(* PLC project Claude3.project, CODESYS CODESYS V3.5 SP20 *)
(* stored: creationDateTime 2026-10-23T09:23:11.8560198, modificationDateTime 2026-10-23T09:22:48.4769723 *)

(* values of E_LineState: DISABLED: Linha desabilitada; WAIT_BOTTLE: Aguardando lote / garrafa; CLAMPING: Cilindro travando a garrafa + tara; FILLING: Enchendo; DRIPPING: Gotejamento, válvula fechada; UNCLAMPING: Cilindro liberando a garrafa; DONE: Ciclo concluído, aguarda avanço da esteira; FAULT: Falha travada, requer reset *)

{attribute 'qualified_only'}
{attribute 'strict'}
TYPE E_LineState : (DISABLED := 0, WAIT_BOTTLE := 1, CLAMPING := 2, FILLING := 3, DRIPPING := 4, UNCLAMPING := 5, DONE := 6, FAULT := 7);
END_TYPE

(* values of E_Fault: FILL_TIMEOUT: Tempo de enchimento excedido; CLAMP_TIMEOUT: Cilindro nao fechou no tempo; UNCLAMP_TIMEOUT: Cilindro nao abriu no tempo; BOTTLE_REMOVED: Garrafa removida durante o ciclo; SAFETY: Emergencia ou porta aberta *)

{attribute 'qualified_only'}
{attribute 'strict'}
TYPE E_Fault : (NONE := 0, FILL_TIMEOUT := 1, CLAMP_TIMEOUT := 2, UNCLAMP_TIMEOUT := 3, BOTTLE_REMOVED := 4, SAFETY := 5);
END_TYPE

(* values of E_ConvState: ADVANCE: Esteira avancando ate o proximo lote; SETTLE: Lote posicionado, tempo de acomodacao; PROCESSING: Linhas enchendo *)

{attribute 'qualified_only'}
{attribute 'strict'}
TYPE E_ConvState : (ADVANCE := 0, SETTLE := 1, PROCESSING := 2);
END_TYPE

TYPE ST_Recipe : STRUCT
  sName : STRING(20);  (* Nome da receita *)
  rTargetMass_g : REAL;  (* Massa liquida alvo [g] *)
  rPreAct_g : REAL;  (* Pre-atuacao: fecha a valvula antes do alvo [g] *)
  rTolerance_g : REAL;  (* Tolerancia +/- para aprovar a garrafa [g] *)
  tFillTimeout : TIME;  (* Tempo maximo de enchimento *)
  tDrip : TIME;  (* Tempo de gotejamento *)
END_STRUCT;
END_TYPE

FUNCTION_BLOCK FB_MovingAvg
  VAR_INPUT
    rIn : REAL;  (* Amostra atual *)
  END_VAR
  VAR_OUTPUT
    rOut : REAL;  (* Media das ultimas C_FILTER_SIZE amostras *)
  END_VAR
  VAR
    aBuf : ARRAY[0..(GVL_Main.C_FILTER_SIZE - 1)] OF REAL;
    iIdx : INT := 0;
    bInit : BOOL := FALSE;
    i : INT;
    rSum : REAL;
  END_VAR

                  (* Na primeira chamada, preenche o buffer para evitar transitorio *)
IF NOT bInit THEN
    FOR i := 0 TO GVL_Main.C_FILTER_SIZE - 1 DO
        aBuf[i] := rIn;
    END_FOR;
    bInit := TRUE;
END_IF;

(* Buffer circular *)
aBuf[iIdx] := rIn;
iIdx := iIdx + 1;
IF iIdx > GVL_Main.C_FILTER_SIZE - 1 THEN
    iIdx := 0;
END_IF;

(* Soma e media *)
rSum := 0.0;
FOR i := 0 TO GVL_Main.C_FILTER_SIZE - 1 DO
    rSum := rSum + aBuf[i];
END_FOR;
rOut := rSum / INT_TO_REAL(GVL_Main.C_FILTER_SIZE);
                
END_FUNCTION_BLOCK

FUNCTION_BLOCK FB_LevelControl
  VAR_INPUT
    bEnable : BOOL;  (* FALSE = fecha a valvula (seguranca) *)
    rLevel_pct : REAL;  (* Nivel atual [%] *)
    rLowOn_pct : REAL := 30.0;  (* Abre a valvula abaixo deste nivel *)
    rHighOff_pct : REAL := 80.0;  (* Fecha a valvula acima deste nivel *)
    rMinOperate_pct : REAL := 15.0;  (* Minimo para liberar o enchimento *)
  END_VAR
  VAR_OUTPUT
    bFillValve : BOOL;  (* Valvula de entrada do tanque *)
    bTankOk : BOOL;  (* Nivel suficiente para envasar *)
    bLowLevelAlarm : BOOL;
  END_VAR

                  (* Histerese: a saida mantem o ultimo estado entre os limites *)
IF NOT bEnable THEN
    bFillValve := FALSE;
ELSIF rLevel_pct <= rLowOn_pct THEN
    bFillValve := TRUE;
ELSIF rLevel_pct >= rHighOff_pct THEN
    bFillValve := FALSE;
END_IF;

(* Permissivo de envase e alarme de nivel baixo *)
bTankOk        := rLevel_pct >= rMinOperate_pct;
bLowLevelAlarm := NOT bTankOk;
                
END_FUNCTION_BLOCK

FUNCTION_BLOCK FB_FillLine
  VAR_INPUT
    bEnable : BOOL;  (* Linha habilitada *)
    bSafetyOk : BOOL;  (* Emergencia e porta OK *)
    bRun : BOOL;  (* Maquina em producao (permite iniciar garrafa) *)
    bLotReady : BOOL;  (* Lote posicionado e acomodado *)
    bTankOk : BOOL;  (* Nivel do tanque suficiente *)
    bBottlePresent : BOOL;
    bClampClosed : BOOL;
    bClampOpen : BOOL;
    bReset : BOOL;  (* Reset de falha (borda de subida) *)
    rMass_g : REAL;  (* Massa bruta filtrada *)
    stRecipe : ST_Recipe;
  END_VAR
  VAR_OUTPUT
    bClampCmd : BOOL;
    bFillValve : BOOL;
    bFinished : BOOL;  (* Desabilitada ou concluida no lote atual *)
    bBusy : BOOL;  (* Garrafa em processo *)
    bFault : BOOL;
    eState : E_LineState := E_LineState.DISABLED;
    eFault : E_Fault := E_Fault.NONE;
    rNetMass_g : REAL;
    diFilled : DINT;
    diRejected : DINT;
  END_VAR
  VAR
    trigReset : R_TRIG;
    tonClamp : TON;
    tonUnclamp : TON;
    tonTare : TON;
    tonFill : TON;
    tonDrip : TON;
    tonBottle : TON;
    rTare_g : REAL;
    bInProcess : BOOL;  (* Ha garrafa em processo nesta linha *)
    bFaultMidCycle : BOOL;  (* Falha ocorreu com garrafa em processo *)
    bWatchBottle : BOOL;
    eFaultNew : E_Fault;
  END_VAR

                  (* ---- 1. Temporizadores e deteccao de borda ---- *)
bWatchBottle := (eState = E_LineState.CLAMPING) OR (eState = E_LineState.FILLING)
                OR (eState = E_LineState.DRIPPING);

trigReset(CLK := bReset);
tonClamp  (IN := (eState = E_LineState.CLAMPING)   AND NOT bClampClosed, PT := GVL_Main.C_T_CYL_TIMEOUT);
tonTare   (IN := (eState = E_LineState.CLAMPING)   AND bClampClosed,     PT := GVL_Main.C_T_TARE);
tonUnclamp(IN := (eState = E_LineState.UNCLAMPING) AND NOT bClampOpen,   PT := GVL_Main.C_T_CYL_TIMEOUT);
tonFill   (IN := (eState = E_LineState.FILLING),                         PT := stRecipe.tFillTimeout);
tonDrip   (IN := (eState = E_LineState.DRIPPING),                        PT := stRecipe.tDrip);
tonBottle (IN := bWatchBottle AND NOT bBottlePresent,                    PT := GVL_Main.C_T_BOTTLE_DEB);

(* ---- 2. Deteccao de falhas (seguranca tem a maior prioridade) ---- *)
eFaultNew := E_Fault.NONE;
IF NOT bSafetyOk THEN
    eFaultNew := E_Fault.SAFETY;
ELSIF tonClamp.Q THEN
    eFaultNew := E_Fault.CLAMP_TIMEOUT;
ELSIF tonUnclamp.Q THEN
    eFaultNew := E_Fault.UNCLAMP_TIMEOUT;
ELSIF tonFill.Q THEN
    eFaultNew := E_Fault.FILL_TIMEOUT;
ELSIF tonBottle.Q THEN
    eFaultNew := E_Fault.BOTTLE_REMOVED;
END_IF;

IF (eFaultNew <> E_Fault.NONE) AND (eState <> E_LineState.FAULT)
   AND (eState <> E_LineState.DISABLED) THEN
    IF bInProcess THEN
        diRejected     := diRejected + 1;     (* Garrafa abortada = rejeitada *)
        bInProcess     := FALSE;
        bFaultMidCycle := TRUE;
    ELSE
        bFaultMidCycle := FALSE;
    END_IF;
    eFault := eFaultNew;
    eState := E_LineState.FAULT;
END_IF;

(* ---- 3. Massa liquida ---- *)
IF (eState = E_LineState.FILLING) OR (eState = E_LineState.DRIPPING) THEN
    rNetMass_g := rMass_g - rTare_g;
ELSIF eState = E_LineState.WAIT_BOTTLE THEN
    rNetMass_g := 0.0;
END_IF;

(* ---- 4. Maquina de estados ---- *)
CASE eState OF

    E_LineState.DISABLED:
        bClampCmd  := FALSE;
        bFillValve := FALSE;
        IF bEnable THEN
            eState := E_LineState.WAIT_BOTTLE;
        END_IF;

    E_LineState.WAIT_BOTTLE:
        bClampCmd  := FALSE;
        bFillValve := FALSE;
        IF NOT bEnable THEN
            eState := E_LineState.DISABLED;
        ELSIF bLotReady AND NOT bBottlePresent THEN
            eState := E_LineState.DONE;                  (* Posicao vazia: nada a envasar *)
        ELSIF bRun AND bLotReady AND bBottlePresent AND bTankOk THEN
            bInProcess := TRUE;
            eState     := E_LineState.CLAMPING;
        END_IF;

    E_LineState.CLAMPING:
        bClampCmd  := TRUE;
        bFillValve := FALSE;
        IF tonTare.Q THEN                                (* Cilindro fechado e massa estavel *)
            rTare_g := rMass_g;
            eState  := E_LineState.FILLING;
        END_IF;

    E_LineState.FILLING:
        bClampCmd := TRUE;
        IF rNetMass_g >= (stRecipe.rTargetMass_g - stRecipe.rPreAct_g) THEN
            bFillValve := FALSE;
            eState     := E_LineState.DRIPPING;
        ELSE
            bFillValve := TRUE;
        END_IF;

    E_LineState.DRIPPING:
        bClampCmd  := TRUE;
        bFillValve := FALSE;
        IF tonDrip.Q THEN
            IF ABS(rNetMass_g - stRecipe.rTargetMass_g) <= stRecipe.rTolerance_g THEN
                diFilled   := diFilled + 1;
            ELSE
                diRejected := diRejected + 1;
            END_IF;
            bInProcess := FALSE;
            eState     := E_LineState.UNCLAMPING;
        END_IF;

    E_LineState.UNCLAMPING:
        bClampCmd  := FALSE;
        bFillValve := FALSE;
        IF bClampOpen THEN
            eState := E_LineState.DONE;
        END_IF;

    E_LineState.DONE:
        bClampCmd  := FALSE;
        bFillValve := FALSE;
        IF NOT bLotReady THEN                            (* Lote saiu: prepara o proximo *)
            IF bEnable THEN
                eState := E_LineState.WAIT_BOTTLE;
            ELSE
                eState := E_LineState.DISABLED;
            END_IF;
        END_IF;

    E_LineState.FAULT:
        bClampCmd  := FALSE;                             (* Valvula fechada e garrafa liberada *)
        bFillValve := FALSE;
        IF trigReset.Q AND bSafetyOk THEN
            eFault := E_Fault.NONE;
            IF bFaultMidCycle THEN
                eState := E_LineState.DONE;              (* Garrafa ja contabilizada como rejeitada *)
            ELSE
                eState := E_LineState.WAIT_BOTTLE;
            END_IF;
            bFaultMidCycle := FALSE;
        END_IF;

END_CASE;

(* ---- 5. Saidas de status ---- *)
bFault    := (eState = E_LineState.FAULT);
bFinished := (eState = E_LineState.DISABLED) OR (eState = E_LineState.DONE);
bBusy     := (eState = E_LineState.CLAMPING) OR (eState = E_LineState.FILLING)
             OR (eState = E_LineState.DRIPPING) OR (eState = E_LineState.UNCLAMPING);
                

METHOD M_ClearCounters : BOOL
                        (* Zera os contadores de garrafas envasadas e rejeitadas da linha *)
diFilled   := 0;
diRejected := 0;
                      
END_METHOD
END_FUNCTION_BLOCK

PROGRAM PRG_Main
  VAR
    aLoadAvg : ARRAY[1..GVL_Main.C_NUM_LINES] OF FB_MovingAvg;
    aLine : ARRAY[1..GVL_Main.C_NUM_LINES] OF FB_FillLine;
    fbTank : FB_LevelControl;
    eConv : E_ConvState := E_ConvState.ADVANCE;
    trigStart : R_TRIG;
    trigLot : R_TRIG;
    tonSettle : TON;
    bSafetyOk : BOOL;  (* Cadeia de seguranca lida pelo CLP; a protecao fisica deve ser independente *)
    bAllFinished : BOOL;
    bAnyFault : BOOL;
    bAnyBusy : BOOL;
    bConvStarted : BOOL;  (* Esteira ja se moveu desde a partida *)
    diSumFilled : DINT;
    diSumRejected : DINT;
    i : INT;
  END_VAR

                  (* ---- 1. Seguranca: emergencia e porta (contatos NF) ---- *)
bSafetyOk := GVL_Main.bEStopOk AND GVL_Main.bGuardClosed;

(* ---- 2. Tanque pulmao com histerese ---- *)
GVL_Main.rTankLevel_pct := FC_Scale(iRaw    := GVL_Main.iTankLevelRaw,
                                    iRawMin := GVL_Main.C_RAW_MIN,
                                    iRawMax := GVL_Main.C_RAW_MAX,
                                    rEngMin := 0.0,
                                    rEngMax := GVL_Main.rTankLevelMax_pct);
fbTank(bEnable         := bSafetyOk,
       rLevel_pct      := GVL_Main.rTankLevel_pct,
       rLowOn_pct      := GVL_Main.rTankLowOn_pct,
       rHighOff_pct    := GVL_Main.rTankHighOff_pct,
       rMinOperate_pct := GVL_Main.rTankMinOperate_pct);
GVL_Main.qTankInletValve := fbTank.bFillValve;

(* ---- 3. Selecao de receita: somente com a maquina parada e sem garrafa em processo ---- *)
GVL_Main.bRecipeLocked := GVL_Main.bRunning OR bAnyBusy;
IF NOT GVL_Main.bRecipeLocked
   AND (GVL_Main.iRecipeReq >= 1) AND (GVL_Main.iRecipeReq <= 3)
   AND (GVL_Main.iRecipeReq <> GVL_Main.iRecipeActive) THEN
    GVL_Main.stActiveRecipe := GVL_Main.aRecipes[GVL_Main.iRecipeReq];
    GVL_Main.iRecipeActive  := GVL_Main.iRecipeReq;
END_IF;

(* ---- 4. Linhas de enchimento ---- *)
bAllFinished  := TRUE;
bAnyFault     := FALSE;
bAnyBusy      := FALSE;
diSumFilled   := 0;
diSumRejected := 0;

FOR i := 1 TO GVL_Main.C_NUM_LINES DO

    (* Escalonamento e media movel da celula de carga *)
    aLoadAvg[i](rIn := FC_Scale(iRaw    := GVL_Main.aiLoadCellRaw[i],
                                iRawMin := GVL_Main.C_RAW_MIN,
                                iRawMax := GVL_Main.C_RAW_MAX,
                                rEngMin := 0.0,
                                rEngMax := GVL_Main.rLoadCellFullScale_g));
    GVL_Main.arMassGross_g[i] := aLoadAvg[i].rOut;

    (* Ciclo da linha *)
    aLine[i](bEnable        := GVL_Main.abLineEnable[i],
             bSafetyOk      := bSafetyOk,
             bRun           := GVL_Main.bRunning,
             bLotReady      := (eConv = E_ConvState.PROCESSING),
             bTankOk        := fbTank.bTankOk,
             bBottlePresent := GVL_Main.abBottlePresent[i],
             bClampClosed   := GVL_Main.abClampClosed[i],
             bClampOpen     := GVL_Main.abClampOpen[i],
             bReset         := GVL_Main.bResetPB,
             rMass_g        := aLoadAvg[i].rOut,
             stRecipe       := GVL_Main.stActiveRecipe);

    (* Zeragem de contadores (pulso) *)
    IF GVL_Main.bClearCounters THEN
        aLine[i].M_ClearCounters();
    END_IF;

    (* Saidas fisicas e diagnostico *)
    GVL_Main.abClampCmd[i]  := aLine[i].bClampCmd;
    GVL_Main.abFillValve[i] := aLine[i].bFillValve;
    GVL_Main.arMassNet_g[i] := aLine[i].rNetMass_g;
    GVL_Main.aeLineState[i] := aLine[i].eState;
    GVL_Main.aeLineFault[i] := aLine[i].eFault;
    GVL_Main.adiFilled[i]   := aLine[i].diFilled;
    GVL_Main.adiRejected[i] := aLine[i].diRejected;

    (* Agregacao *)
    IF NOT aLine[i].bFinished THEN
        bAllFinished := FALSE;
    END_IF;
    IF aLine[i].bFault THEN
        bAnyFault := TRUE;
    END_IF;
    IF aLine[i].bBusy THEN
        bAnyBusy := TRUE;
    END_IF;
    diSumFilled   := diSumFilled   + aLine[i].diFilled;
    diSumRejected := diSumRejected + aLine[i].diRejected;

END_FOR;

GVL_Main.bClearCounters   := FALSE;
GVL_Main.diTotalFilled    := diSumFilled;
GVL_Main.diTotalRejected  := diSumRejected;

(* ---- 5. Liga/desliga da maquina ---- *)
trigStart(CLK := GVL_Main.bStartPB);
IF (NOT bSafetyOk) OR bAnyFault OR GVL_Main.bStopPB THEN
    GVL_Main.bRunning := FALSE;                          (* Emergencia/porta/falha/parada *)
ELSIF trigStart.Q AND (GVL_Main.iRecipeActive >= 1) THEN
    GVL_Main.bRunning := TRUE;
END_IF;

(* ---- 6. Sequenciamento da esteira ---- *)
trigLot(CLK := GVL_Main.bLotInPos);
tonSettle(IN := (eConv = E_ConvState.SETTLE) AND GVL_Main.bRunning,
          PT := GVL_Main.C_T_SETTLE);

CASE eConv OF

    E_ConvState.ADVANCE:
        (* Borda de subida do sensor = novo lote; na 1a partida aceita lote ja posicionado *)
        IF trigLot.Q
           OR (GVL_Main.bLotInPos AND NOT bConvStarted AND GVL_Main.bRunning) THEN
            eConv := E_ConvState.SETTLE;
        END_IF;

    E_ConvState.SETTLE:
        IF tonSettle.Q THEN
            eConv := E_ConvState.PROCESSING;
        END_IF;

    E_ConvState.PROCESSING:
        (* Todas as linhas habilitadas concluidas: avanca o proximo lote *)
        IF bAllFinished AND GVL_Main.bRunning THEN
            bConvStarted := TRUE;
            eConv        := E_ConvState.ADVANCE;
        END_IF;

END_CASE;

GVL_Main.qConveyor := GVL_Main.bRunning AND bSafetyOk AND (eConv = E_ConvState.ADVANCE);

(* ---- 7. Alarmes ---- *)
GVL_Main.bAlarmAny  := bAnyFault OR fbTank.bLowLevelAlarm;
GVL_Main.qAlarmLamp := GVL_Main.bAlarmAny;
                
END_PROGRAM

FUNCTION FC_Scale : REAL
  VAR_INPUT
    iRaw : INT;  (* Valor bruto do canal analogico *)
    iRawMin : INT;  (* Bruto minimo (0) *)
    iRawMax : INT;  (* Bruto maximo (27648) *)
    rEngMin : REAL;  (* Engenharia no bruto minimo *)
    rEngMax : REAL;  (* Engenharia no bruto maximo *)
  END_VAR
  VAR
    rX : REAL;
  END_VAR

                  (* Protecao contra divisao por zero *)
IF iRawMax = iRawMin THEN
    FC_Scale := rEngMin;
    RETURN;
END_IF;

(* Limita o bruto a faixa valida *)
rX := LIMIT(INT_TO_REAL(iRawMin), INT_TO_REAL(iRaw), INT_TO_REAL(iRawMax));

(* Interpolacao linear *)
FC_Scale := rEngMin + (rX - INT_TO_REAL(iRawMin)) * (rEngMax - rEngMin)
            / (INT_TO_REAL(iRawMax) - INT_TO_REAL(iRawMin));
                
END_FUNCTION

CONFIGURATION Application
  RESOURCE Application ON PLC
    {attribute 'qualified_only'}
    VAR_GLOBAL CONSTANT  (* GVL_Main *)
      C_NUM_LINES : INT := 4;
      C_FILTER_SIZE : INT := 10;  (* Amostras da media movel *)
      C_RAW_MIN : INT := 0;
      C_RAW_MAX : INT := 27648;
      C_T_CYL_TIMEOUT : TIME := TIME#2s0ms;  (* Tempo maximo de movimento do cilindro *)
      C_T_BOTTLE_DEB : TIME := TIME#300ms;  (* Filtro da garrafa removida *)
      C_T_TARE : TIME := TIME#1s0ms;  (* Estabilizacao antes da tara *)
      C_T_SETTLE : TIME := TIME#500ms;  (* Acomodacao do lote *)
      aiLoadCellRaw AT %IW0 : ARRAY[1..4] OF INT;  (* Celulas de carga 1..4 *)
      iTankLevelRaw AT %IW8 : INT;  (* Nivel do tanque *)
      abBottlePresent AT %IX0.0 : ARRAY[1..4] OF BOOL;  (* Sensor de garrafa *)
      abClampClosed AT %IX1.0 : ARRAY[1..4] OF BOOL;  (* Cilindro recuado/travado *)
      abClampOpen AT %IX2.0 : ARRAY[1..4] OF BOOL;  (* Cilindro liberado *)
      bEStopOk AT %IX3.0 : BOOL;  (* TRUE = emergencia rearmada (NF) *)
      bGuardClosed AT %IX3.1 : BOOL;  (* TRUE = porta fechada (NF) *)
      bLotInPos AT %IX3.2 : BOOL;  (* Lote posicionado *)
      bStartPB AT %IX3.3 : BOOL;  (* Botao liga (NA) *)
      bStopPB AT %IX3.4 : BOOL;  (* Botao desliga (NA) *)
      bResetPB AT %IX3.5 : BOOL;  (* Botao reset de falhas (NA) *)
      abClampCmd AT %QX0.0 : ARRAY[1..4] OF BOOL;  (* TRUE = travar garrafa *)
      abFillValve AT %QX1.0 : ARRAY[1..4] OF BOOL;  (* TRUE = valvula aberta *)
      qConveyor AT %QX2.0 : BOOL;
      qTankInletValve AT %QX2.1 : BOOL;
      qAlarmLamp AT %QX2.2 : BOOL;
      rLoadCellFullScale_g : REAL := 1000.0;  (* Massa correspondente a 27648 [g] *)
      rTankLevelMax_pct : REAL := 100.0;
      rTankLowOn_pct : REAL := 30.0;  (* Liga reposicao *)
      rTankHighOff_pct : REAL := 80.0;  (* Desliga reposicao *)
      rTankMinOperate_pct : REAL := 15.0;  (* Minimo para iniciar enchimento *)
      abLineEnable : ARRAY[1..4] OF BOOL := [4(TRUE)];  (* ---- Interface com IHM ---- *)
      aRecipes : ARRAY[1..3] OF ST_Recipe := [(sName := 'Receita 1', rTargetMass_g := 250.0, rPreAct_g := 4.0, rTolerance_g := 3.0, tFillTimeout := TIME#10s0ms, tDrip := TIME#1s0ms), (sName := 'Receita 2', rTargetMass_g := 500.0, rPreAct_g := 6.0, rTolerance_g := 4.0, tFillTimeout := TIME#15s0ms, tDrip := TIME#1s500ms), (sName := 'Receita 3', rTargetMass_g := 750.0, rPreAct_g := 8.0, rTolerance_g := 5.0, tFillTimeout := TIME#20s0ms, tDrip := TIME#2s0ms)];
      iRecipeReq : INT := 1;  (* Receita solicitada (1..3) *)
      iRecipeActive : INT := 0;  (* Receita em uso *)
      stActiveRecipe : ST_Recipe;
      bRecipeLocked : BOOL;  (* TRUE = troca de receita bloqueada *)
      bClearCounters : BOOL;  (* Zera contadores (pulso) *)
      bRunning : BOOL;  (* ---- Estado e diagnostico ---- *)
      bAlarmAny : BOOL;
      rTankLevel_pct : REAL;
      arMassGross_g : ARRAY[1..4] OF REAL;
      arMassNet_g : ARRAY[1..4] OF REAL;
      aeLineState : ARRAY[1..4] OF E_LineState;
      aeLineFault : ARRAY[1..4] OF E_Fault;
      adiFilled : ARRAY[1..4] OF DINT;
      adiRejected : ARRAY[1..4] OF DINT;
      diTotalFilled : DINT;
      diTotalRejected : DINT;
    END_VAR
    TASK MainTask(INTERVAL := T#20ms, PRIORITY := 1);
    PROGRAM PRG_Main WITH MainTask : PRG_Main;
    PROGRAM PLC_PRG WITH MainTask : PLC_PRG;
  END_RESOURCE
END_CONFIGURATION
